// TIA Portal V21 export
// export: Created 2026-10-12T11:32:13.6401694Z, ExportSetting WithDefaults, DisplayName Totally Integrated Automation Portal, DisplayVersion V21, DisplayName STEP 7 Professional, DisplayVersion V21, DisplayName STEP 7 Safety, DisplayVersion V21, DisplayName Tech WebApplication, DisplayVersion V21, DisplayName WinCC Basic/Comfort/Advanced, DisplayVersion V21, DisplayName WinCC Unified, DisplayVersion V21
FUNCTION "FC_GENERAL" : Void   // FC1, LAD
{ S7_Optimized_Access := 'TRUE' }
VERSION : 0.1
// stored: AutoNumber true, IsIECCheckEnabled false, SetENOAutomatically false, UDAEnableTagReadback false
BEGIN

REGION Network 1: CONTROL ON
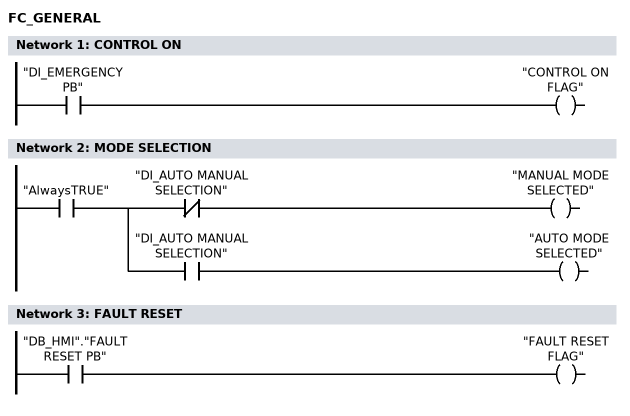
   RUNG wire#powerrail
      Contact( "DI_EMERGENCY PB" )
      Coil( "CONTROL ON FLAG" )
   END_RUNG
   // the same network as SCL:
   "CONTROL ON FLAG" := "DI_EMERGENCY PB";
END_REGION

REGION Network 2: MODE SELECTION
   RUNG wire#powerrail
      Contact( "AlwaysTRUE" )
      wire#w1
      I_Contact( "DI_AUTO MANUAL SELECTION" )
      Coil( "MANUAL MODE SELECTED" )
   END_RUNG
   RUNG wire#w1
      Contact( "DI_AUTO MANUAL SELECTION" )
      Coil( "AUTO MODE SELECTED" )
   END_RUNG
   // the same network as SCL:
   "MANUAL MODE SELECTED" := "AlwaysTRUE" AND NOT "DI_AUTO MANUAL SELECTION";
   "AUTO MODE SELECTED" := "AlwaysTRUE" AND "DI_AUTO MANUAL SELECTION";
END_REGION

REGION Network 3: FAULT RESET
   RUNG wire#powerrail
      Contact( "DB_HMI"."FAULT RESET PB" )
      Coil( "FAULT RESET FLAG" )
   END_RUNG
   // the same network as SCL:
   "FAULT RESET FLAG" := "DB_HMI"."FAULT RESET PB";
END_REGION
END_FUNCTION
